FUNCTION_BLOCK MagazineSupplyWp (* Basic Function Block Type *)
  (* Standard: 61499-2 *)
  (* Version 0.0, 7/2/2026, Template *)
  PACKAGE Main;
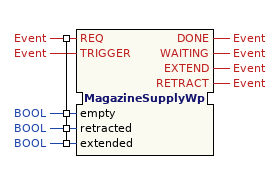
  EVENT_INPUT
    REQ WITH empty, retracted, extended; (* Normal Execution Request *)
    TRIGGER;
  END_EVENT
  EVENT_OUTPUT
    DONE;
    WAITING;
    EXTEND;
    RETRACT;
  END_EVENT
  VAR_INPUT
    empty : BOOL; (* Input event qualifier *)
    retracted : BOOL;
    extended : BOOL;
  END_VAR
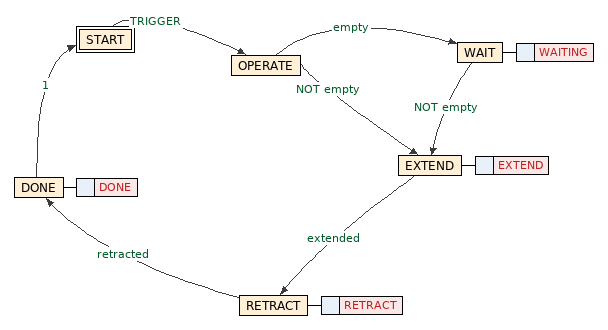
  EC_STATES
    START; (* Initial State *)
    OPERATE;
    EXTEND : -> EXTEND;
    RETRACT : -> RETRACT;
    DONE : -> DONE;
    WAIT : -> WAITING;
  END_STATES
  EC_TRANSITIONS
    DONE TO START := 1;
    START TO OPERATE := TRIGGER;
    OPERATE TO EXTEND := NOT empty;
    OPERATE TO WAIT := empty;
    WAIT TO EXTEND := NOT empty;
    EXTEND TO RETRACT := extended;
    RETRACT TO DONE := retracted;
  END_TRANSITIONS
  ALGORITHM INIT IN ST: (* Initialization algorithm *)
;
  END_ALGORITHM
  ALGORITHM REQ IN ST: (* Normally executed algorithm *)
;
  END_ALGORITHM
END_FUNCTION_BLOCK
